// TIA Portal V21 export
DATA_BLOCK "IDB_SclSections"   // DB4
// stored: InstanceOfName FB_SclSections, InstanceOfType FB
"FB_SclSections"
   // VAR_INPUT
   //    Enable : Bool := TRUE;
   //    Mode : Int := 2;
   //    Setpoint : Real := 50.0;
   // END_VAR
   // VAR_OUTPUT
   //    Busy : Bool := TRUE;
   //    Result : Real;
   //    StepCount : Int;
   // END_VAR
   // VAR_IN_OUT
   //    Values : Array[0..9] of Real;
   // END_VAR
   // VAR
   //    State : Int := 10;
   //    Sum : Real := 12.5;
   //    Iterations : Int := 3;
   // END_VAR
BEGIN
END_DATA_BLOCK
